(* IEC 61131-3 sources: iolistgen/tests_support/pl_stub/src/DUTs/AnalogInput, 8 files *)

(* ---- E_AiAlarm.dut.st ---- *)
// Назначение: заглушка plc-process-lib 1.0.0 для проверки типов сгенерированного кода без CODESYS
//             (API.md, раздел 4.1); не библиотека — тел и внутренних переменных нет
// Автор:      kr0nsch
// Версия:     1.0.0 (выпуск библиотеки)
// Документ:   docs/GENERATORS.md, раздел «Проверка ST без CODESYS»
{attribute 'qualified_only'}
TYPE E_AiAlarm :
(
    HH := 0,
    H := 1,
    L := 2,
    LL := 3,
    Failure := 4,
    OutOfRange := 5
) UINT;
END_TYPE

(* ---- E_AiFailValue.dut.st ---- *)
// Назначение: заглушка plc-process-lib 1.0.0 для проверки типов сгенерированного кода без CODESYS
//             (API.md, раздел 11.1); не библиотека — тел и внутренних переменных нет
// Автор:      kr0nsch
// Версия:     1.0.0 (выпуск библиотеки)
// Документ:   docs/GENERATORS.md, раздел «Проверка ST без CODESYS»
{attribute 'qualified_only'}
{attribute 'strict'}
TYPE E_AiFailValue :
(
    HoldLast := 0,
    Substitute := 1
) INT;
END_TYPE

(* ---- E_AiInputType.dut.st ---- *)
// Назначение: заглушка plc-process-lib 1.0.0 для проверки типов сгенерированного кода без CODESYS
//             (API.md, раздел 11.1); не библиотека — тел и внутренних переменных нет
// Автор:      kr0nsch
// Версия:     1.0.0 (выпуск библиотеки)
// Документ:   docs/GENERATORS.md, раздел «Проверка ST без CODESYS»
{attribute 'qualified_only'}
{attribute 'strict'}
TYPE E_AiInputType :
(
    MilliAmp := 0,
    Norm420 := 1,
    Norm01 := 2,
    Eng := 3,
    Raw := 4
) INT;
END_TYPE

(* ---- E_AiSignalState.dut.st ---- *)
// Назначение: заглушка plc-process-lib 1.0.0 для проверки типов сгенерированного кода без CODESYS
//             (API.md, раздел 11.1); не библиотека — тел и внутренних переменных нет
// Автор:      kr0nsch
// Версия:     1.0.0 (выпуск библиотеки)
// Документ:   docs/GENERATORS.md, раздел «Проверка ST без CODESYS»
{attribute 'qualified_only'}
{attribute 'strict'}
TYPE E_AiSignalState :
(
    Good := 0,
    UnderRange := 1,
    OverRange := 2,
    FailLow := 3,
    FailHigh := 4,
    ChannelFault := 5,
    NotFinite := 6
) INT;
END_TYPE

(* ---- ST_AiLimitCfg.dut.st ---- *)
// Назначение: заглушка plc-process-lib 1.0.0 для проверки типов сгенерированного кода без CODESYS
//             (API.md, раздел 8.3); не библиотека — тел и внутренних переменных нет
// Автор:      kr0nsch
// Версия:     1.0.0 (выпуск библиотеки)
// Документ:   docs/GENERATORS.md, раздел «Проверка ST без CODESYS»
{attribute 'qualified_only'}
TYPE ST_AiLimitCfg :
STRUCT
    xEnable      : BOOL := FALSE;
    rSetpoint_eu : REAL := 0.0;
    rHyst_eu     : REAL := 0.0;
    tOnDelay     : TIME := T#0S;
    tOffDelay    : TIME := T#0S;
END_STRUCT
END_TYPE

(* ---- ST_AnalogInputCfg.dut.st ---- *)
// Назначение: заглушка plc-process-lib 1.0.0 для проверки типов сгенерированного кода без CODESYS
//             (API.md, раздел 11.1); не библиотека — тел и внутренних переменных нет
// Автор:      kr0nsch
// Версия:     1.0.0 (выпуск библиотеки)
// Документ:   docs/GENERATORS.md, раздел «Проверка ST без CODESYS»
{attribute 'qualified_only'}
TYPE ST_AnalogInputCfg :
STRUCT
    eInput         : E_AiInputType := E_AiInputType.MilliAmp;
    rRangeLo_eu    : REAL := 0.0;
    rRangeHi_eu    : REAL := 100.0;
    rRawLo_cnt     : REAL := 0.0;
    rRawHi_cnt     : REAL := 0.0;
    xSqrt          : BOOL := FALSE;
    rLowCut_pct    : REAL := 0.0;
    tFilter        : TIME := T#0S;
    tFailDelay     : TIME := T#2S;
    eFailValue     : E_AiFailValue := E_AiFailValue.HoldLast;
    rFailValue_eu  : REAL := 0.0;
    xLimitsOnFail  : BOOL := FALSE;
    xClamp         : BOOL := FALSE;
    // lint:allow STL007 имя массива по контракту API.md (префикс a + тип элемента)
    astLimit       : ARRAY[0..3] OF ST_AiLimitCfg;
    tSubstMax      : TIME := T#8H;
    udiAlarmIdBase : UDINT := 0;
    // lint:allow STL007 имя массива по контракту API.md (префикс a + тип элемента)
    astAlarm       : ARRAY[0..GVL_Const.DEV_ALARMS_MAX - 1] OF ST_AlarmCfg := [
            (ePriority := E_AlarmPriority.High),
            (ePriority := E_AlarmPriority.Low),
            (ePriority := E_AlarmPriority.Low),
            (ePriority := E_AlarmPriority.High),
            (ePriority := E_AlarmPriority.Medium),
            (ePriority := E_AlarmPriority.Low),
            (ePriority := E_AlarmPriority.None),
            (ePriority := E_AlarmPriority.None)];
END_STRUCT
END_TYPE

(* ---- ST_AnalogInputCmd.dut.st ---- *)
// Назначение: заглушка plc-process-lib 1.0.0 для проверки типов сгенерированного кода без CODESYS
//             (API.md, раздел 11.1); не библиотека — тел и внутренних переменных нет
// Автор:      kr0nsch
// Версия:     1.0.0 (выпуск библиотеки)
// Документ:   docs/GENERATORS.md, раздел «Проверка ST без CODESYS»
{attribute 'qualified_only'}
TYPE ST_AnalogInputCmd :
STRUCT
    stCommon       : ST_DeviceCmd;
    rSubstValue_eu : REAL;
END_STRUCT
END_TYPE

(* ---- ST_AnalogInputSts.dut.st ---- *)
// Назначение: заглушка plc-process-lib 1.0.0 для проверки типов сгенерированного кода без CODESYS
//             (API.md, раздел 11.1); не библиотека — тел и внутренних переменных нет
// Автор:      kr0nsch
// Версия:     1.0.0 (выпуск библиотеки)
// Документ:   docs/GENERATORS.md, раздел «Проверка ST без CODESYS»
{attribute 'qualified_only'}
TYPE ST_AnalogInputSts :
STRUCT
    stCommon        : ST_DeviceSts;
    rValue_eu       : REAL;
    rValue_pct      : REAL;
    rIn             : REAL;
    eSignal         : E_AiSignalState;
    uiSubstRemain_s : UINT;
END_STRUCT
END_TYPE
